// Mock of the mirror covers. A subclass of HalfBROT.FB_CoverControl, since FB_MonetTelescopeControl takes the concrete block (it calls
// Stop(), which I_MirrorCovers does not carry); the real body (limit switches, AT%I*/AT%Q*, timers) does not run (no SUPER^()), as for
// the axis mocks. With nMockTravelScans = 0 (default) Open/Close take effect at once. With nMockTravelScans > 0 a run takes that many
// calls of the body (FB_MonetRig.Scan calls it after the telescope, the MAIN order): Open()/Close() latch the direction as the real
// block does and Stop() drops it, so the covers stay where they are (neither Opened nor Closed in between). After InjectError() the
// covers report an error and do not move (HalfBROT FB_CoverControl inhibits every cover output while bError), until Reset();
// Open/Close/Stop are still counted.
FUNCTION_BLOCK FB_CoversMock EXTENDS HalfBROT.FB_CoverControl
VAR_INPUT
	nMockTravelScans	: UINT;	// scans a full open or close takes, 0 = at once (FB_MonetRig.SetCoverTravelScans)
END_VAR
VAR
	bOpened		: BOOL;
	bClosed		: BOOL := TRUE;
	bFailed		: BOOL;
	nOpenCalls	: UINT;
	nCloseCalls	: UINT;
	nStopCalls	: UINT;
	bRunOpen	: BOOL;	// an open runs (nMockTravelScans > 0)
	bRunClose	: BOOL;	// a close runs
	nTravelPos	: UINT;	// 0 = closed .. nMockTravelScans = open
END_VAR

// No SUPER^(): only the travel model below runs
IF bFailed THEN
	bRunOpen := FALSE;
	bRunClose := FALSE;
ELSIF bRunOpen THEN
	IF nTravelPos < nMockTravelScans THEN
		nTravelPos := nTravelPos + 1;
	END_IF
	IF nTravelPos >= nMockTravelScans THEN
		bRunOpen := FALSE;
	END_IF
ELSIF bRunClose THEN
	IF nTravelPos > 0 THEN
		nTravelPos := nTravelPos - 1;
	END_IF
	IF nTravelPos = 0 THEN
		bRunClose := FALSE;
	END_IF
END_IF
IF nMockTravelScans > 0 THEN
	bOpened := nTravelPos >= nMockTravelScans;
	bClosed := nTravelPos = 0;
END_IF
bAllOpen := bOpened;
bAllClosed := bClosed;
bError := bFailed;

METHOD Open : BOOL
IF NOT bFailed THEN
	IF nMockTravelScans = 0 THEN
		bOpened := TRUE;
		bClosed := FALSE;
	ELSE
		bRunOpen := TRUE;
		bRunClose := FALSE;
	END_IF
END_IF
nOpenCalls := nOpenCalls + 1;
Open := NOT bFailed;
END_METHOD

METHOD Close : BOOL
IF NOT bFailed THEN
	IF nMockTravelScans = 0 THEN
		bOpened := FALSE;
		bClosed := TRUE;
		nTravelPos := 0;
	ELSE
		bRunClose := TRUE;
		bRunOpen := FALSE;
	END_IF
END_IF
nCloseCalls := nCloseCalls + 1;
Close := NOT bFailed;
END_METHOD

// drops a running open or close: the covers stay where they are (HalfBROT FB_CoverControl.Stop)
METHOD Stop : BOOL
bRunOpen := FALSE;
bRunClose := FALSE;
nStopCalls := nStopCalls + 1;
Stop := TRUE;
END_METHOD

// the covers report an error (Error) and stop where they are until Reset() (MonetSafeState_Tests)
METHOD InjectError
bFailed := TRUE;
END_METHOD

METHOD Reset : BOOL
bFailed := FALSE;
Reset := TRUE;
END_METHOD

PROPERTY Opened : BOOL
GET
Opened := bOpened;
END_GET
END_PROPERTY

PROPERTY Closed : BOOL
GET
Closed := bClosed;
END_GET
END_PROPERTY

PROPERTY Error : BOOL
GET
Error := bFailed;
END_GET
END_PROPERTY

END_FUNCTION_BLOCK

(* stored: Version 1.1.0.1, ProductVersion 3.1.4024.15
   POU FB_CoversMock: Id {f17dfb05-8c2f-48a0-9523-e0aa4e3eb81e}, SpecialFunc None
   Method Open: Id {878b5598-7bb7-4d16-819f-f7ff964312ca}
   Method Close: Id {dc54c13f-ffe1-4494-9ce6-0a5905cb5ccc}
   Method Stop: Id {c4becc20-75cd-4a2b-9be2-342968dc4e3a}
   Method InjectError: Id {63619404-82d7-479d-8d28-e715d56d9cfa}
   Method Reset: Id {0b918468-8437-4bae-bedb-9b7a9531322e}
   Property Opened: Id {9f0d87fc-b2be-4fac-a4ec-8deb394287bf}
   Get Get: Id {53e0617a-fd86-42b6-a811-84d49e77466b}
   Property Closed: Id {ffcda306-0a5f-43bd-936b-bffbde33e1c0}
   Get Get: Id {0aef944c-4a5c-471f-9558-f7beefc93bc4}
   Property Error: Id {ccafefc7-a111-4388-91b0-2dd3fd487173}
   Get Get: Id {23c63bde-cc9b-40e4-b598-8aa868f352a3} *)
